SUBAPPLICATION OptionalGroup_001b (* Optionsgruppe 1b: Digitaler Eingang/Ausgang per Options-Adapter freigeschaltet (QI aus AOption_X_TO_EVENT aktiviert/deaktiviert die ganze Gruppe) - letztes Glied einer Daisy-Chain, reicht nichts weiter. *)
  (* Standard: 61499-2; Description: Copyright (c) 2026 Meisterschulen am Ostbahnhof This program and the accompanying materials are made available under the terms of the Eclipse Public License 2.0 which is available at https://www.eclipse.org/legal/epl-2.0/ SPDX-License-Identifier: EPL-2.0 *)
  (* Version 1.0, 2026-10-13, Franz Höpfinger, Meisterschulen am Ostbahnhof, Baugleich zu OptionalGroup_001a, aber ohne PLUG1 - wird typischerweise an PLUG1 einer vorgeschalteten OptionalGroup_001a angehaengt, damit beide Gruppen nacheinander (erst a, dann b) aktiviert werden, bevor der urspruengliche Aufrufer seine Bestaetigung erhaelt. *)
  PACKAGE MyLib_AX_Option::sys;
  IMPORT logiBUS::io::DI::logiBUS_DI::Input_I1;
  IMPORT logiBUS::io::DQ::logiBUS_DO::Output_Q1;
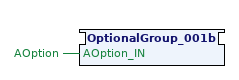
  SOCKETS
    AOption_IN : Option::AOption;
  END_SOCKETS
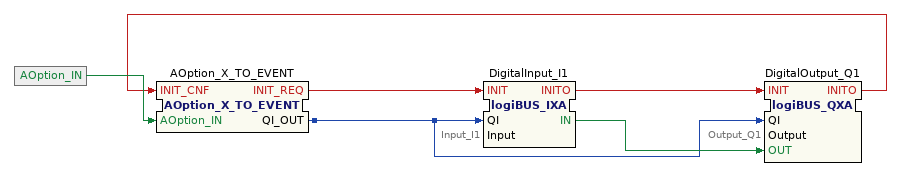
  FBS
    DigitalInput_I1 : logiBUS::io::DI::logiBUS_IXA(Input := Input_I1);
    DigitalOutput_Q1 : logiBUS::io::DQ::logiBUS_QXA(Output := Output_Q1);
    AOption_X_TO_EVENT : Option::conversion::AOption_X_TO_EVENT;
  END_FBS
  EVENT_CONNECTIONS
    AOption_X_TO_EVENT.INIT_REQ TO DigitalInput_I1.INIT;
    DigitalInput_I1.INITO TO DigitalOutput_Q1.INIT;
    DigitalOutput_Q1.INITO TO AOption_X_TO_EVENT.INIT_CNF;
  END_CONNECTIONS
  DATA_CONNECTIONS
    AOption_X_TO_EVENT.QI_OUT TO DigitalInput_I1.QI;
    AOption_X_TO_EVENT.QI_OUT TO DigitalOutput_Q1.QI;
  END_CONNECTIONS
  ADAPTER_CONNECTIONS
    DigitalInput_I1.IN TO DigitalOutput_Q1.OUT;
    AOption_IN TO AOption_X_TO_EVENT.AOption_IN;
  END_CONNECTIONS
END_SUBAPPLICATION
